Staubli VAL3: action.dtx

public num nActResult
public num nActType
public num nActIO
